FUNCTION_BLOCK Gradeamento_Inovaisa_HMI (* Service Interface Function Block Type *)
  (* Standard: 61499-2 *)
  (* Version 1.0, 22/10/2026, Hidryco, Hidryco, IHM do Gradeamento_Inovaisa *)
  PACKAGE Hidryco.HidrycoLib;
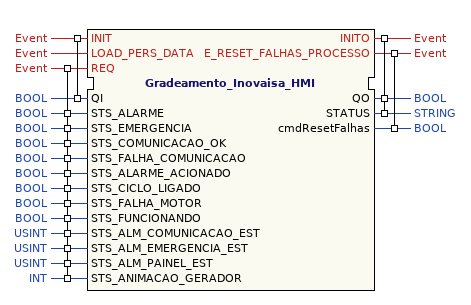
  EVENT_INPUT
    INIT WITH QI;
    LOAD_PERS_DATA; (* Reenvia os parametros persistentes *)
    REQ WITH STS_ALARME, STS_EMERGENCIA, STS_COMUNICACAO_OK, STS_FALHA_COMUNICACAO, STS_ALARME_ACIONADO, STS_CICLO_LIGADO, STS_FALHA_MOTOR, STS_FUNCIONANDO, STS_ALM_COMUNICACAO_EST, STS_ALM_EMERGENCIA_EST, STS_ALM_PAINEL_EST, STS_ANIMACAO_GERADOR; (* Atualizacao de status *)
  END_EVENT
  EVENT_OUTPUT
    INITO WITH QO, STATUS;
    E_RESET_FALHAS_PROCESSO WITH cmdResetFalhas;
  END_EVENT
  VAR_INPUT
    QI : BOOL;
    STS_ALARME : BOOL; (* Algum alarme do gradeamento (comunicacao, painel, emergencia, motores) *)
    STS_EMERGENCIA : BOOL; (* Botao de emergencia do painel acionado (4006) *)
    STS_COMUNICACAO_OK : BOOL; (* Comunicacao Modbus com o CLP do painel OK *)
    STS_FALHA_COMUNICACAO : BOOL; (* Falha de comunicacao com o CLP do painel *)
    STS_ALARME_ACIONADO : BOOL; (* Alarme acionado no painel (4005) *)
    STS_CICLO_LIGADO : BOOL; (* Comando de ciclo remoto ligado (4001 = 1) *)
    STS_FALHA_MOTOR : BOOL; (* Grade ou rosca em falha ou sobretorque *)
    STS_FUNCIONANDO : BOOL; (* Alguma grade ou a rosca funcionando *)
    STS_ALM_COMUNICACAO_EST : USINT; (* Estado do ALARM_BIT (0 normal, 1 ativo reconhecido, 2 ativo nao reconhecido, 3 saiu nao reconhecido, 4 ativo e saiu nao reconhecido) *)
    STS_ALM_EMERGENCIA_EST : USINT; (* Estado do ALARM_BIT (0 normal, 1 ativo reconhecido, 2 ativo nao reconhecido, 3 saiu nao reconhecido, 4 ativo e saiu nao reconhecido) *)
    STS_ALM_PAINEL_EST : USINT; (* Estado do ALARM_BIT (0 normal, 1 ativo reconhecido, 2 ativo nao reconhecido, 3 saiu nao reconhecido, 4 ativo e saiu nao reconhecido) *)
    STS_ANIMACAO_GERADOR : INT; (* Raio do gerador: 0 nao conectado, 1 nao liberada, 2 liberada, 3 liberada e funcionando nos geradores *)
  END_VAR
  VAR_OUTPUT
    QO : BOOL; (* Event Output Qualifier *)
    STATUS : STRING; (* Service Status *)
    cmdResetFalhas : BOOL; (* Reset do painel (4002), dos sensores e reconhecimento dos alarmes do gradeamento *)
  END_VAR
  SERVICE /
    SEQUENCE 
    END_SEQUENCE
  END_SERVICE
END_FUNCTION_BLOCK
